Fanuc KAREL source: KB00056.KL

PROGRAM KB00056
%NOLOCKGROUP
VAR
  P1: INTEGER
  P2: BOOLEAN
  P3: INTEGER
BEGIN
  P1 = 1
  P2 = TRUE
  P3 = 1
  DAQ_STOP(P1, P2, P3)
END KB00056
